Staubli VAL3: main.pgx

program main()
begin
  close(tCurrentTool)
  pPointRx.config.shoulder = lefty
  pPointRx.config.elbow = epositive
  pPointRx.config.wrist = wpositive
  pPointRx2.config.shoulder = lefty
  pPointRx2.config.elbow = epositive
  pPointRx2.config.wrist = wpositive
  mCurrentSpeed.tvel = 100.00
  mCurrentSpeed.blend = joint
  mCurrentSpeed.reach = 0.010
  mCurrentSpeed.leave = 0.010
  // Program TgtProg start
  // Program generated by RoboDK v6.0.7 for Staubli RX130B on XX/XX/XXXX 18:00:00
  // Using nominal kinematics.
  Output[1]=true
  Output[1]=false
  Output[1]=true
  Output[1]=x
  Output[1]=true
  Output[2]=false
  Output[2]=y
  Output[2]=true
  watch(Input[1]==true)
  watch(Input[1]==false)
  watch(Input[1]==x)
  watch(Input[1]==true,0.0)
  watch(V==true,1234.6)
  V=false

  waitEndMove()
  // Program TgtProg end

end
